(* IEC 61131-3 sources: llm-plc-st-eval/data/processed_definitivo/gpt-4o-2024-08-06/B6/zero_shot, 3 files *)

(* ---- ejec_1.st ---- *)
FUNCTION_BLOCK FB_Baliza
VAR_INPUT
    alarma : BOOL; // Variable de entrada que indica si hay una condición de alarma
END_VAR

VAR_OUTPUT
    lampara : BOOL; // Variable de salida que controla el estado de la lámpara
END_VAR

VAR
    temporizador : TON; // Temporizador para controlar el parpadeo
    estado_parpadeo : BOOL; // Estado interno para el parpadeo
END_VAR

// Inicialización del temporizador
temporizador(IN := estado_parpadeo, PT := T#1S);

// Lógica de control de la baliza
IF alarma THEN
    temporizador(IN := NOT temporizador.Q); // Alterna el estado del temporizador
    estado_parpadeo := temporizador.Q; // Actualiza el estado de parpadeo
    lampara := estado_parpadeo; // La lámpara sigue el estado de parpadeo
ELSE
    temporizador(IN := FALSE); // Resetea el temporizador si no hay alarma
    estado_parpadeo := FALSE; // Asegura que el estado de parpadeo esté apagado
    lampara := FALSE; // Apaga la lámpara si no hay alarma
END_IF
END_FUNCTION_BLOCK

(* ---- ejec_2.st ---- *)
FUNCTION_BLOCK FB_Baliza
VAR_INPUT
    alarma : BOOL; // Variable de entrada que indica si hay una condición de alarma
END_VAR

VAR_OUTPUT
    lampara : BOOL; // Variable de salida que controla el estado de la lámpara
END_VAR

VAR
    temporizador : TON; // Temporizador para controlar el parpadeo
    estado_parpadeo : BOOL; // Estado interno para alternar el parpadeo
END_VAR

// Inicialización del temporizador
temporizador(IN := estado_parpadeo, PT := T#1S);

IF alarma THEN
    // Si hay alarma, activar el temporizador
    temporizador(IN := NOT temporizador.Q);

    // Alternar el estado de parpadeo cuando el temporizador termina
    IF temporizador.Q THEN
        estado_parpadeo := NOT estado_parpadeo;
    END_IF;

    // La lámpara sigue el estado de parpadeo
    lampara := estado_parpadeo;
ELSE
    // Si no hay alarma, apagar la lámpara y reiniciar el temporizador
    lampara := FALSE;
    estado_parpadeo := FALSE;
    temporizador(IN := FALSE);
END_IF;

END_FUNCTION_BLOCK

(* ---- ejec_3.st ---- *)
FUNCTION_BLOCK FB_Baliza
VAR_INPUT
    alarma : BOOL; // Entrada que indica si hay una condición de alarma
END_VAR

VAR_OUTPUT
    lampara : BOOL; // Salida que controla el estado de la lámpara
END_VAR

VAR
    timerBlink : TON; // Temporizador para el parpadeo de la lámpara
    estadoParpadeo : BOOL; // Estado interno para el parpadeo
END_VAR

// Inicialización del temporizador
timerBlink(IN := estadoParpadeo, PT := T#1S);

// Lógica de control de la baliza
IF alarma THEN
    // Si hay alarma, alternar el estado de parpadeo cada segundo
    IF timerBlink.Q THEN
        estadoParpadeo := NOT estadoParpadeo;
        timerBlink(IN := FALSE); // Reiniciar el temporizador
    ELSE
        timerBlink(IN := TRUE); // Activar el temporizador
    END_IF;
    lampara := estadoParpadeo; // Actualizar el estado de la lámpara
ELSE
    // Si no hay alarma, la lámpara está apagada
    lampara := FALSE;
    estadoParpadeo := FALSE; // Reiniciar el estado de parpadeo
    timerBlink(IN := FALSE); // Asegurarse de que el temporizador esté desactivado
END_IF;
END_FUNCTION_BLOCK
